// TIA Portal V20 export
Screen "Barcode_Scanner"  1276x673
  ScreenItem "线_1" at 0,81 size 1366x2  Type=HmiLine
  ScreenItem "permanentareaborderrectangle" at 0,0 size 0x0  Type=HmiRectangle
  ScreenItem "Button_Back" at 3,12 size 90x60  Type=HmiButton
  ScreenItem "Title_OPMode1_ScreenOverview_X390_Y2" at 433,7 size 500x30  Type=HmiTextBox
  ScreenItem "符号 IO 域_1" at 451,38 size 475x42  Type=HmiSymbolicIOField
